Fanuc KAREL source: kc00027.KL

-- PROVISIONAL review KL for V940-1; original PC SHA256 748457f7056725b1c834b0ef74314b3c5bba6a6d14d1efada8d8826d942d761e
-- Incomplete behavior may be omitted. Consult companion uncertainty JSON. Do not deploy.
PROGRAM KC00027
%NOLOCKGROUP
BEGIN
  -- V9_ZERO_TABLE_METADATA_HINT layout=0002_ascii; no indexed target words; source/name/runtime held
  -- UNRESOLVED_PC offsets 5-81; opcodes 27,22,1C,22,1C,22,1C,22,22,1C,22,22,22,31
  -- UNRESOLVED_PC offsets 86-90; opcodes 7F
END KC00027
